Staubli VAL3: utText.pjx

--- utText.pjx ---
Parameters version=s8.10Cs9_BS1925 stackSize=5000 millimeterUnit=true
Program file=start.pgx
Program file=stop.pgx
Data file=utText.dtx
Type name=utCommon path=./utCommon/utCommon.pjx
Type name=utText path=./utText/utText.pjx
Type name=utBorder path=./utBorder/utBorder.pjx
Type name=utAppearance path=./utAppearance/utAppearance.pjx

--- utText.dtx ---
public utCommon Common
  [0]
    bool bDisabled
    string sValue
    string sID
    num nValue
    string sPage
public utText Text
  [0]
    string sFontFamily
    string sFontStyle
    string sFontWeight
    string sTextAlignment
    num nFontSize
public utBorder Border
  [0]
    string sBorderColour
    string sBorderSytle
    string sBorderWidth
public utAppearance Appearance
  [0]
    string sBackgroundColour
    string sColour
    bool bVisibility

--- start.pgx ---
program start()
begin
end

--- stop.pgx ---
program stop()
begin
end
